ADAPTER system_info (* Adapter Interface *)
  (* Standard: 61499-1 *)
  (* Version 0.0, 10/23/2026, macie, Schneider Electric *)
  PACKAGE Main;
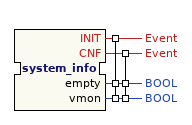
  EVENT_OUTPUT
    INIT WITH vmon, empty;
    CNF WITH vmon, empty; (* Confirmation from Plug *)
  END_EVENT
  VAR_OUTPUT
    empty : BOOL; (* Indication Data from Plug *)
    vmon : BOOL; (* Confirmation Data from Plug *)
  END_VAR
  SERVICE SOCKET/PLUG
    SEQUENCE request_confirm
      SOCKET.REQ(REQD) -> PLUG.REQ(REQD);
      PLUG.CNF(vmon) -> SOCKET.CNF(vmon);
    END_SEQUENCE
    SEQUENCE indication_response
      PLUG.IND(empty) -> SOCKET.IND(empty);
      SOCKET.RSP(RSPD) -> PLUG.RSP(RSPD);
    END_SEQUENCE
  END_SERVICE
END_ADAPTER
